(* PLC project GeneratedProgram, SafePLC-Gen SafePLC-Gen Multimodal 1.0 *)
(* stored: creationDateTime 2026-04-25T13:53:54.159190Z *)

PROGRAM GeneratedProgram
  VAR
    LOOP_4750_03_TRIP : BOOL;
    LOOP_4712_02_TRIP : BOOL;
    LOOP_104_01_TRIP : BOOL;
    TICSA_4750_03_HH : BOOL;
    TICSA_4750_03_LL : BOOL;
    PICSA_4712_02_HH : BOOL;
    PICSA_4712_02_LL : BOOL;
    SV_104_01_HH : BOOL;
    SV_104_01_LL : BOOL;
    SAFE_STATE : BOOL;
    FirstScan : BOOL;
    TICSA_4750_03_Scaled : REAL;
    PICSA_4712_02_Scaled : REAL;
    PI_4712_01_Scaled : REAL;
    TICSA_4750_03_HH_SP : REAL;
    TICSA_4750_03_H_SP : REAL;
    TICSA_4750_03_L_SP : REAL;
    TICSA_4750_03_LL_SP : REAL;
    TICSA_4750_03_Deadband : REAL;
    PICSA_4712_02_HH_SP : REAL;
    PICSA_4712_02_H_SP : REAL;
    PICSA_4712_02_L_SP : REAL;
    PICSA_4712_02_LL_SP : REAL;
    PICSA_4712_02_Deadband : REAL;
    PI_4712_01_HH_SP : REAL;
    PI_4712_01_H_SP : REAL;
    PI_4712_01_L_SP : REAL;
    PI_4712_01_LL_SP : REAL;
    PI_4712_01_Deadband : REAL;
    TICSA_4750_03_H : BOOL;
    TICSA_4750_03_L : BOOL;
    TICSA_4750_03_HH_Latch : SR;
    TICSA_4750_03_LL_Latch : SR;
    TICSA_4750_03_HH_Ack : BOOL;
    TICSA_4750_03_LL_Ack : BOOL;
    PICSA_4712_02_H : BOOL;
    PICSA_4712_02_L : BOOL;
    PICSA_4712_02_HH_Latch : SR;
    PICSA_4712_02_LL_Latch : SR;
    PICSA_4712_02_HH_Ack : BOOL;
    PICSA_4712_02_LL_Ack : BOOL;
    PI_4712_01_H : BOOL;
    PI_4712_01_L : BOOL;
    PI_4712_01_HH_Latch : SR;
    PI_4712_01_LL_Latch : SR;
    PI_4712_01_HH_Ack : BOOL;
    PI_4712_01_LL_Ack : BOOL;
    TICSA_4750_03_SP : REAL;
    TICSA_4750_03_Kp : REAL;
    TICSA_4750_03_Ki : REAL;
    TICSA_4750_03_Integral : REAL;
    TICSA_4750_03_Error : REAL;
    TICSA_4750_03_Output_Pct : REAL;
    PICSA_4712_02_SP : REAL;
    PICSA_4712_02_Kp : REAL;
    PICSA_4712_02_Ki : REAL;
    PICSA_4712_02_Integral : REAL;
    PICSA_4712_02_Error : REAL;
    PICSA_4712_02_Output_Pct : REAL;
    XV_HS_4750_01_Cmd : BOOL;
    System_Alarm : BOOL;
  END_VAR

            IF FirstScan THEN
    LOOP_4750_03_TRIP := TRUE;
    LOOP_4712_02_TRIP := TRUE;
    LOOP_104_01_TRIP  := TRUE;
    SAFE_STATE        := TRUE;
    TV_4750_03_Out    := 32767;
    PVA_4712_02_Out   := 6554;
    MV_MNb_47121_Out  := 6554;
    MV_MNb_47122_Out  := 6554;
    MV_MNb_47123_Out  := 6554;
    MV_MNc_47124_Out  := 6554;
    MV_MNc_47125a_Out := 6554;
    MV_MNc_47125b_Out := 6554;
    MV_MNc_47126_Out  := 6554;
    MV_MNc_47127_Out  := 6554;
    MV_WKa_47130_Out  := 6554;
    MV_WKa_47131_Out  := 6554;
    MV_73KH12_50a_Out := 6554;
    MV_73KH12_50b_Out := 6554;
    MV_73KH12_50c_Out := 6554;
    MV_73KH12_25_Out  := 6554;
    MV_QSa_47140_Out  := 6554;
    MV_QSb_47141_Out  := 6554;
    XV_HS_4750_01     := FALSE;
    FirstScan         := FALSE;
    RETURN;
END_IF;

TICSA_4750_03_Scaled := ((INT_TO_REAL(TICSA_4750_03_Raw) - 6554.0) / (32767.0 - 6554.0)) * 200.0;
PICSA_4712_02_Scaled := ((INT_TO_REAL(PICSA_4712_02_Raw) - 6554.0) / (32767.0 - 6554.0)) * 100.0;
PI_4712_01_Scaled    := ((INT_TO_REAL(PI_4712_01_Raw)    - 6554.0) / (32767.0 - 6554.0)) * 100.0;

IF TICSA_4750_03_Scaled >= TICSA_4750_03_HH_SP THEN
    TICSA_4750_03_HH := TRUE;
ELSIF TICSA_4750_03_Scaled <= (TICSA_4750_03_HH_SP - TICSA_4750_03_Deadband) THEN
    TICSA_4750_03_HH := FALSE;
END_IF;

IF TICSA_4750_03_Scaled >= TICSA_4750_03_H_SP THEN
    TICSA_4750_03_H := TRUE;
ELSIF TICSA_4750_03_Scaled <= (TICSA_4750_03_H_SP - TICSA_4750_03_Deadband) THEN
    TICSA_4750_03_H := FALSE;
END_IF;

IF TICSA_4750_03_Scaled <= TICSA_4750_03_LL_SP THEN
    TICSA_4750_03_LL := TRUE;
ELSIF TICSA_4750_03_Scaled >= (TICSA_4750_03_LL_SP + TICSA_4750_03_Deadband) THEN
    TICSA_4750_03_LL := FALSE;
END_IF;

IF TICSA_4750_03_Scaled <= TICSA_4750_03_L_SP THEN
    TICSA_4750_03_L := TRUE;
ELSIF TICSA_4750_03_Scaled >= (TICSA_4750_03_L_SP + TICSA_4750_03_Deadband) THEN
    TICSA_4750_03_L := FALSE;
END_IF;

TICSA_4750_03_HH_Latch(S1 := TICSA_4750_03_HH,
                        R  := (TICSA_4750_03_HH_Ack AND NOT TICSA_4750_03_HH));
TICSA_4750_03_LL_Latch(S1 := TICSA_4750_03_LL,
                        R  := (TICSA_4750_03_LL_Ack AND NOT TICSA_4750_03_LL));

IF PICSA_4712_02_Scaled >= PICSA_4712_02_HH_SP THEN
    PICSA_4712_02_HH := TRUE;
ELSIF PICSA_4712_02_Scaled <= (PICSA_4712_02_HH_SP - PICSA_4712_02_Deadband) THEN
    PICSA_4712_02_HH := FALSE;
END_IF;

IF PICSA_4712_02_Scaled >= PICSA_4712_02_H_SP THEN
    PICSA_4712_02_H := TRUE;
ELSIF PICSA_4712_02_Scaled <= (PICSA_4712_02_H_SP - PICSA_4712_02_Deadband) THEN
    PICSA_4712_02_H := FALSE;
END_IF;

IF PICSA_4712_02_Scaled <= PICSA_4712_02_LL_SP THEN
    PICSA_4712_02_LL := TRUE;
ELSIF PICSA_4712_02_Scaled >= (PICSA_4712_02_LL_SP + PICSA_4712_02_Deadband) THEN
    PICSA_4712_02_LL := FALSE;
END_IF;

IF PICSA_4712_02_Scaled <= PICSA_4712_02_L_SP THEN
    PICSA_4712_02_L := TRUE;
ELSIF PICSA_4712_02_Scaled >= (PICSA_4712_02_L_SP + PICSA_4712_02_Deadband) THEN
    PICSA_4712_02_L := FALSE;
END_IF;

PICSA_4712_02_HH_Latch(S1 := PICSA_4712_02_HH,
                        R  := (PICSA_4712_02_HH_Ack AND NOT PICSA_4712_02_HH));
PICSA_4712_02_LL_Latch(S1 := PICSA_4712_02_LL,
                        R  := (PICSA_4712_02_LL_Ack AND NOT PICSA_4712_02_LL));

IF PI_4712_01_Scaled >= PI_4712_01_HH_SP THEN
    PI_4712_01_HH_Latch(S1 := TRUE, R := FALSE);
ELSIF PI_4712_01_Scaled <= (PI_4712_01_HH_SP - PI_4712_01_Deadband) THEN
    PI_4712_01_HH_Latch(S1 := FALSE, R := (PI_4712_01_HH_Ack AND NOT (PI_4712_01_Scaled >= PI_4712_01_HH_SP)));
END_IF;

IF PI_4712_01_Scaled >= PI_4712_01_H_SP THEN
    PI_4712_01_H := TRUE;
ELSIF PI_4712_01_Scaled <= (PI_4712_01_H_SP - PI_4712_01_Deadband) THEN
    PI_4712_01_H := FALSE;
END_IF;

IF PI_4712_01_Scaled <= PI_4712_01_LL_SP THEN
    PI_4712_01_LL_Latch(S1 := TRUE, R := FALSE);
ELSIF PI_4712_01_Scaled >= (PI_4712_01_LL_SP + PI_4712_01_Deadband) THEN
    PI_4712_01_LL_Latch(S1 := FALSE, R := (PI_4712_01_LL_Ack AND NOT (PI_4712_01_Scaled <= PI_4712_01_LL_SP)));
END_IF;

IF PI_4712_01_Scaled <= PI_4712_01_L_SP THEN
    PI_4712_01_L := TRUE;
ELSIF PI_4712_01_Scaled >= (PI_4712_01_L_SP + PI_4712_01_Deadband) THEN
    PI_4712_01_L := FALSE;
END_IF;

IF TICSA_4750_03_HH OR TICSA_4750_03_LL THEN
    LOOP_4750_03_TRIP := TRUE;
ELSIF LOOP_4750_03_TRIP AND MANUAL_RESET
      AND NOT TICSA_4750_03_HH AND NOT TICSA_4750_03_LL THEN
    LOOP_4750_03_TRIP := FALSE;
END_IF;

IF PICSA_4712_02_HH OR PICSA_4712_02_LL THEN
    LOOP_4712_02_TRIP := TRUE;
ELSIF LOOP_4712_02_TRIP AND MANUAL_RESET
      AND NOT PICSA_4712_02_HH AND NOT PICSA_4712_02_LL THEN
    LOOP_4712_02_TRIP := FALSE;
END_IF;

IF SV_104_01_HH OR SV_104_01_LL THEN
    LOOP_104_01_TRIP := TRUE;
ELSIF LOOP_104_01_TRIP AND MANUAL_RESET
      AND NOT SV_104_01_HH AND NOT SV_104_01_LL THEN
    LOOP_104_01_TRIP := FALSE;
END_IF;

SAFE_STATE := ESTOP OR LOOP_4750_03_TRIP OR LOOP_4712_02_TRIP OR LOOP_104_01_TRIP;

IF NOT SAFE_STATE THEN
    XV_HS_4750_01_Cmd := HS_4750_01;
    XV_HS_4750_01     := XV_HS_4750_01_Cmd;
ELSE
    XV_HS_4750_01_Cmd := FALSE;
    XV_HS_4750_01     := FALSE;
END_IF;

IF NOT SAFE_STATE THEN
    TICSA_4750_03_Error    := TICSA_4750_03_SP - TICSA_4750_03_Scaled;
    TICSA_4750_03_Integral := TICSA_4750_03_Integral + (TICSA_4750_03_Ki * TICSA_4750_03_Error);
    IF TICSA_4750_03_Integral > 100.0 THEN
        TICSA_4750_03_Integral := 100.0;
    ELSIF TICSA_4750_03_Integral < 0.0 THEN
        TICSA_4750_03_Integral := 0.0;
    END_IF;
    TICSA_4750_03_Output_Pct := (TICSA_4750_03_Kp * TICSA_4750_03_Error) + TICSA_4750_03_Integral;
    IF TICSA_4750_03_Output_Pct > 100.0 THEN
        TICSA_4750_03_Output_Pct := 100.0;
    ELSIF TICSA_4750_03_Output_Pct < 0.0 THEN
        TICSA_4750_03_Output_Pct := 0.0;
    END_IF;
    TV_4750_03_Out := REAL_TO_INT(6554.0 + (TICSA_4750_03_Output_Pct / 100.0) * (32767.0 - 6554.0));
ELSE
    TV_4750_03_Out := 32767;
END_IF;

IF NOT SAFE_STATE THEN
    PICSA_4712_02_Error    := PICSA_4712_02_SP - PICSA_4712_02_Scaled;
    PICSA_4712_02_Integral := PICSA_4712_02_Integral + (PICSA_4712_02_Ki * PICSA_4712_02_Error);
    IF PICSA_4712_02_Integral > 100.0 THEN
        PICSA_4712_02_Integral := 100.0;
    ELSIF PICSA_4712_02_Integral < 0.0 THEN
        PICSA_4712_02_Integral := 0.0;
    END_IF;
    PICSA_4712_02_Output_Pct := (PICSA_4712_02_Kp * PICSA_4712_02_Error) + PICSA_4712_02_Integral;
    IF PICSA_4712_02_Output_Pct > 100.0 THEN
        PICSA_4712_02_Output_Pct := 100.0;
    ELSIF PICSA_4712_02_Output_Pct < 0.0 THEN
        PICSA_4712_02_Output_Pct := 0.0;
    END_IF;
    PVA_4712_02_Out := REAL_TO_INT(6554.0 + (PICSA_4712_02_Output_Pct / 100.0) * (32767.0 - 6554.0));
ELSE
    PVA_4712_02_Out := 6554;
END_IF;

IF SAFE_STATE THEN
    MV_MNb_47121_Out  := 6554;
    MV_MNb_47122_Out  := 6554;
    MV_MNb_47123_Out  := 6554;
    MV_MNc_47124_Out  := 6554;
    MV_MNc_47125a_Out := 6554;
    MV_MNc_47125b_Out := 6554;
    MV_MNc_47126_Out  := 6554;
    MV_MNc_47127_Out  := 6554;
    MV_WKa_47130_Out  := 6554;
    MV_WKa_47131_Out  := 6554;
    MV_73KH12_50a_Out := 6554;
    MV_73KH12_50b_Out := 6554;
    MV_73KH12_50c_Out := 6554;
    MV_73KH12_25_Out  := 6554;
    MV_QSa_47140_Out  := 6554;
    MV_QSb_47141_Out  := 6554;
END_IF;

System_Alarm :=
    TICSA_4750_03_HH_Latch.Q1 OR TICSA_4750_03_LL_Latch.Q1 OR
    TICSA_4750_03_H            OR TICSA_4750_03_L            OR
    PICSA_4712_02_HH_Latch.Q1 OR PICSA_4712_02_LL_Latch.Q1 OR
    PICSA_4712_02_H            OR PICSA_4712_02_L            OR
    PI_4712_01_HH_Latch.Q1    OR PI_4712_01_LL_Latch.Q1    OR
    PI_4712_01_H               OR PI_4712_01_L              OR
    LOOP_4750_03_TRIP          OR LOOP_4712_02_TRIP         OR
    LOOP_104_01_TRIP           OR SAFE_STATE;
          
END_PROGRAM

CONFIGURATION Config0
  RESOURCE Res0 ON PLC
    TASK MainTask(INTERVAL := T#20ms, PRIORITY := 0);
    PROGRAM Main : GeneratedProgram;
  END_RESOURCE
END_CONFIGURATION
